// TIA Portal V20 export
Screen "Pop-up_Opmodes18_Popup"  645x340
  ScreenItem "Background" at 0,0 size 645x339  Type=HmiRectangle
  ScreenItem "Descr_HmiPanel" at 1,283 size 56x40  Type=HmiTextBox
  ScreenItem "Linie1_LightGrey" at 10,282 size 520x0  Type=HmiLine
  ScreenItem "Linie1_DarkGrey" at 10,281 size 520x0  Type=HmiLine
  ScreenItem "Linie1_LightGrey_1" at 10,324 size 520x0  Type=HmiLine
  ScreenItem "Linie1_DarkGrey_1" at 10,323 size 520x0  Type=HmiLine
  ScreenItem "Overview_OPMode" at 1,1 size 643x25  Type=HmiTextBox
  ScreenItem "Descr_OPMode" at 1,26 size 550x40  Type=HmiTextBox
  ScreenItem "OPMode17_small" at 540,136 size 90x60  Type=HmiButton
  ScreenItem "OPMode1_small" at 15,71 size 90x60  Type=HmiButton
  ScreenItem "OPMode2_small" at 15,136 size 90x60  Type=HmiButton
  ScreenItem "OPMode3_small" at 15,202 size 90x60  Type=HmiButton
  ScreenItem "OPMode4_small" at 120,71 size 90x60  Type=HmiButton
  ScreenItem "OPMode7_small" at 225,71 size 90x60  Type=HmiButton
  ScreenItem "OPMode5_small" at 121,136 size 90x60  Type=HmiButton
  ScreenItem "OPMode8_small" at 226,136 size 90x60  Type=HmiButton
  ScreenItem "OPMode10_small" at 330,71 size 90x60  Type=HmiButton
  ScreenItem "OPMode11_small" at 331,136 size 90x60  Type=HmiButton
  ScreenItem "OPMode13_small" at 435,71 size 90x60  Type=HmiButton
  ScreenItem "OPMode14_small" at 435,136 size 90x60  Type=HmiButton
  ScreenItem "OPMode16_small" at 540,71 size 90x60  Type=HmiButton
  ScreenItem "OPMode18_small" at 541,202 size 90x60  Type=HmiButton
  ScreenItem "OPMode6_small" at 122,202 size 90x60  Type=HmiButton
  ScreenItem "OPMode9_small" at 227,202 size 90x60  Type=HmiButton
  ScreenItem "OPMode12_small" at 332,202 size 90x60  Type=HmiButton
  ScreenItem "OPMode15_small" at 436,202 size 90x60  Type=HmiButton
  ScreenItem "OPMode1_wide" at 10,71 size 100x60  Type=HmiButton
  ScreenItem "OPMode2_wide" at 10,136 size 100x60  Type=HmiButton
  ScreenItem "OPMode3_wide" at 10,202 size 100x60  Type=HmiButton
  ScreenItem "OPMode4_wide" at 115,71 size 100x60  Type=HmiButton
  ScreenItem "OPMode5_wide" at 115,136 size 100x60  Type=HmiButton
  ScreenItem "OPMode6_wide" at 115,202 size 100x60  Type=HmiButton
  ScreenItem "OPMode7_wide" at 220,71 size 100x60  Type=HmiButton
  ScreenItem "OPMode8_wide" at 220,136 size 100x60  Type=HmiButton
  ScreenItem "OPMode9_wide" at 220,202 size 100x60  Type=HmiButton
  ScreenItem "OPMode10_wide" at 325,71 size 100x60  Type=HmiButton
  ScreenItem "OPMode11_wide" at 325,136 size 100x60  Type=HmiButton
  ScreenItem "OPMode12_wide" at 325,202 size 100x60  Type=HmiButton
  ScreenItem "OPMode13_wide" at 430,71 size 100x60  Type=HmiButton
  ScreenItem "OPMode14_wide" at 430,136 size 100x60  Type=HmiButton
  ScreenItem "OPMode15_wide" at 430,202 size 100x60  Type=HmiButton
  ScreenItem "OPMode16_wide" at 535,71 size 100x60  Type=HmiButton
  ScreenItem "OPMode17_wide" at 535,136 size 100x60  Type=HmiButton
  ScreenItem "OPMode18_wide" at 535,202 size 100x60  Type=HmiButton
  ScreenItem "Overview_HMI-OP" at 554,275 size 90x60  Type=HmiButton
  ScreenItem "Cancel Mode" at 554,1 size 90x60  Type=HmiButton
  ScreenItem "OPMode1_Foreground_Blocked" at 10,71 size 100x60  Type=HmiGraphicView
  ScreenItem "OPMode2_Foreground_Blocked" at 10,136 size 100x60  Type=HmiGraphicView
  ScreenItem "OPMode3_Foreground_Blocked" at 10,202 size 100x60  Type=HmiGraphicView
  ScreenItem "OPMode4_Foreground_Blocked" at 115,71 size 100x60  Type=HmiGraphicView
  ScreenItem "OPMode5_Foreground_Blocked" at 115,136 size 100x60  Type=HmiGraphicView
  ScreenItem "OPMode6_Foreground_Blocked" at 115,202 size 100x60  Type=HmiGraphicView
  ScreenItem "OPMode7_Foreground_Blocked" at 220,71 size 100x60  Type=HmiGraphicView
  ScreenItem "OPMode8_Foreground_Blocked" at 220,136 size 100x60  Type=HmiGraphicView
  ScreenItem "OPMode9_Foreground_Blocked" at 220,202 size 100x60  Type=HmiGraphicView
  ScreenItem "OPMode10_Foreground_Blocked" at 325,71 size 100x60  Type=HmiGraphicView
  ScreenItem "OPMode11_Foreground_Blocked" at 325,136 size 100x60  Type=HmiGraphicView
  ScreenItem "OPMode12_Foreground_Blocked" at 325,202 size 100x60  Type=HmiGraphicView
  ScreenItem "OPMode13_Foreground_Blocked" at 430,71 size 100x60  Type=HmiGraphicView
  ScreenItem "OPMode14_Foreground_Blocked" at 430,136 size 100x60  Type=HmiGraphicView
  ScreenItem "OPMode15_Foreground_Blocked" at 430,202 size 100x60  Type=HmiGraphicView
  ScreenItem "OPMode16_Foreground_Blocked" at 535,71 size 100x60  Type=HmiGraphicView
  ScreenItem "OPMode17_Foreground_Blocked" at 535,136 size 100x60  Type=HmiGraphicView
  ScreenItem "OPMode18_Foreground_Blocked" at 535,202 size 100x60  Type=HmiGraphicView
  ScreenItem "OPMode1_Blocked" at 95,75 size 14x14  Type=HmiGraphicView
  ScreenItem "OPMode2_Blocked" at 95,140 size 14x14  Type=HmiGraphicView
  ScreenItem "OPMode3_Blocked" at 95,205 size 14x14  Type=HmiGraphicView
  ScreenItem "OPMode4_Blocked" at 200,75 size 14x14  Type=HmiGraphicView
  ScreenItem "OPMode5_Blocked" at 200,140 size 14x14  Type=HmiGraphicView
  ScreenItem "OPMode6_Blocked" at 200,205 size 14x14  Type=HmiGraphicView
  ScreenItem "OPMode7_Blocked" at 305,75 size 14x14  Type=HmiGraphicView
  ScreenItem "OPMode8_Blocked" at 305,140 size 14x14  Type=HmiGraphicView
  ScreenItem "OPMode9_Blocked" at 305,205 size 14x14  Type=HmiGraphicView
  ScreenItem "OPMode10_Blocked" at 410,75 size 14x14  Type=HmiGraphicView
  ScreenItem "OPMode11_Blocked" at 410,140 size 14x14  Type=HmiGraphicView
  ScreenItem "OPMode12_Blocked" at 410,205 size 14x14  Type=HmiGraphicView
  ScreenItem "OPMode13_Blocked" at 515,75 size 14x14  Type=HmiGraphicView
  ScreenItem "OPMode14_Blocked" at 515,140 size 14x14  Type=HmiGraphicView
  ScreenItem "OPMode15_Blocked" at 515,205 size 14x14  Type=HmiGraphicView
  ScreenItem "OPMode16_Blocked" at 620,75 size 14x14  Type=HmiGraphicView
  ScreenItem "OPMode17_Blocked" at 620,140 size 14x14  Type=HmiGraphicView
  ScreenItem "OPMode18_Blocked" at 620,205 size 14x14  Type=HmiGraphicView
